FUNCTION_BLOCK FB_Jog
VAR_INPUT
	JogButton	:	INT;
END_VAR
VAR_OUTPUT
	bBusy		:	BOOL;
	bError		:	BOOL;
END_VAR
VAR_IN_OUT
	mot			:	AXIS_REF;
END_VAR
VAR
	fb_MCJog	:	MC_Jog;
END_VAR

CASE ABS(JogButton) OF
	0:	fb_MCJog(
			Axis	:=	mot);
	1:	fb_MCJog(
			Axis	:=	mot,
			Mode	:=	E_JogMode.MC_JOGMODE_STANDARD_SLOW);
	2:	fb_MCJog(
			Axis	:=	mot,
			Mode	:=	E_JogMode.MC_JOGMODE_STANDARD_FAST);
	3:	fb_MCJog(
			Axis	:=	mot,
			Mode	:=	E_JogMode.MC_JOGMODE_CONTINOUS,
			Velocity:=	STRING_TO_LREAL(UserVar.JogTargVel)/60.0);
END_CASE

IF JogButton > 0 THEN
	fb_MCJog.JogForward	:=	TRUE;
	fb_MCJog.JogBackwards	:=	FALSE;
END_IF

IF JogButton < 0 THEN
	fb_MCJog.JogForward	:=	FALSE;
	fb_MCJog.JogBackwards	:=	TRUE;
END_IF

IF JogButton = 0 THEN
	fb_MCJog.JogForward	:=	FALSE;
	fb_MCJog.JogBackwards	:=	FALSE;
END_IF

bBusy	:=	fb_MCJog.Busy;
bError	:=	fb_MCJog.Error;

END_FUNCTION_BLOCK

(* stored: Version 1.1.0.1, ProductVersion 3.1.4024.15
   POU FB_Jog: Id {7aa4005f-be43-41da-b380-71f88d9e71ed}, SpecialFunc None *)
